FUNCTION_BLOCK CycleCounter (* Basic Function Block Type *)
  (* Standard: 61499-2 *)
  (* Version 0.0, 10/21/2026, Schneider Electric, Template *)
  PACKAGE SE.Nereda;
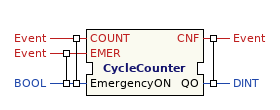
  EVENT_INPUT
    COUNT WITH EmergencyON;
    EMER WITH EmergencyON; (* Normal Execution Request *)
  END_EVENT
  EVENT_OUTPUT
    CNF WITH QO; (* Execution Confirmation *)
  END_EVENT
  VAR_INPUT
    EmergencyON : BOOL; (* Input event qualifier *)
  END_VAR
  VAR_OUTPUT
    QO : DINT; (* Output event qualifier *)
  END_VAR
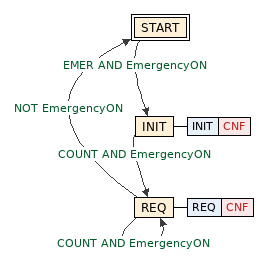
  EC_STATES
    START; (* Initial State *)
    INIT : INIT -> CNF; (* Initialization *)
    REQ : REQ -> CNF; (* Normal execution *)
  END_STATES
  EC_TRANSITIONS
    START TO INIT := EMER AND EmergencyON;
    INIT TO REQ := COUNT AND EmergencyON;
    REQ TO START := NOT EmergencyON;
    REQ TO REQ := COUNT AND EmergencyON;
  END_TRANSITIONS
  ALGORITHM INIT IN ST: (* Initialization algorithm *)
;
QO := 0;
  END_ALGORITHM
  ALGORITHM REQ IN ST: (* Normally executed algorithm *)
;
QO := QO + 1;
COUNT := FALSE;
  END_ALGORITHM
END_FUNCTION_BLOCK
